PROGRAM MAIN
VAR
	// TcUnit finds every FB_TestSuite instance by itself; it is enough to declare them here.
	fbHydraulicsTests	: FB_HydraulicsControl_Tests;
	fbCoverTests		: FB_CoverControl_Tests;
	fbPendantTests		: FB_PendantControl_Tests;
	fbFocusUnlockTests	: FB_FocusUnlock_Tests;
	fbBrakeCloseHoldTests	: FB_BrakeCloseHold_Tests;	// MONETcommon#277
	fbFocusHoldOnStopTests	: F_FocusHoldOnStop_Tests;	// MONETcommon#278
END_VAR

TcUnit.RUN();

END_PROGRAM

(* stored: Version 1.1.0.1, ProductVersion 3.1.4024.15
   POU MAIN: Id {862d57cc-8a35-5254-a921-b66855b6453b}, SpecialFunc None *)
